Fanuc KAREL source: KT00487.KL

PROGRAM KT00487
%NOLOCKGROUP
VAR
  P1: POSITION
  P2: XYZWPREXT
  OUT: JOINTPOS
BEGIN
    P2.Y = 2.0
  OUT = P1 : P2
END KT00487
